// TIA Portal V19 export
TYPE "AnaMon.HMI"
   STRUCT
      identName : String;
      comment : String;
      MsgSupOp : Bool;
      PVScale : Struct
         High : Real := 100.0;
         Low : Real;
      END_STRUCT;
      HiAlmSupOp : Bool;
      HiWrnSupOp : Bool;
      LoWrnSupOp : Bool;
      LoAlmSupOp : Bool;
      PermissionLog { S7_SetPoint := 'True'} : "AnaMon.Permission";
      Status { S7_SetPoint := 'True'} : "AnaMon.Status";
   END_STRUCT;
END_TYPE
